// TIA Portal V20 export
Screen "Dry_runFunction Select"  1225x440
  ScreenItem "Background" at 0,0 size 1221x434  Type=HmiRectangle
  ScreenItem "Overview_Special" at 2,1 size 1219x73  Type=HmiTextBox
  ScreenItem "Faceplate container_1" at 2,77 size 407x119  Type=HmiFaceplateContainer
  ScreenItem "Faceplate container_2" at 407,77 size 406x119  Type=HmiFaceplateContainer
  ScreenItem "Faceplate container_4" at 2,193 size 407x119  Type=HmiFaceplateContainer
  ScreenItem "Faceplate container_7" at 813,77 size 408x119  Type=HmiFaceplateContainer
  ScreenItem "Faceplate container_5" at 408,193 size 408x119  Type=HmiFaceplateContainer
  ScreenItem "Faceplate container_10" at 813,196 size 408x119  Type=HmiFaceplateContainer
  ScreenItem "Faceplate container_11" at 2,313 size 408x119  Type=HmiFaceplateContainer
  ScreenItem "Faceplate container_12" at 407,313 size 408x119  Type=HmiFaceplateContainer
